// TIA Portal V17 export
// export: Created 2026-11-10T15:00:48.6641979Z, ExportSetting WithDefaults, DisplayName Totally Integrated Automation Portal, DisplayVersion V17, DisplayName TIA Portal Openness, DisplayVersion V17, DisplayName TIA Portal Version Control Interface, DisplayVersion V17, DisplayName STEP 7 Professional, DisplayVersion V17, DisplayName STEP 7 Safety, DisplayVersion V17, DisplayName WinCC Advanced, DisplayVersion V17
GraphicList "Lamp_Green"  ListRange=Decimal, Mode=Simple
  GraphicListEntry   EntryType=Range, Picture=Signal_Off
  GraphicListEntry   EntryType=Range, From=1, To=1, Picture=Signal_Green
